FUNCTION_BLOCK ActuatorBaseExt (* Composite Function Block Type *)
  (* Standard: 61499-2 *)
  (* Version 1.0.1, 10/17/2023, ApplicationLibDevTeam, Schneider Electric, First Version *)
  PACKAGE Flexbridge.FestoMPS400;
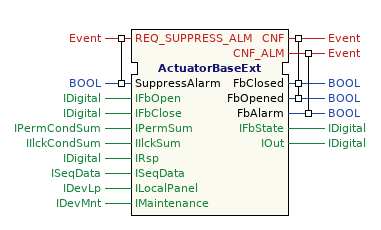
  EVENT_INPUT
    REQ_SUPPRESS_ALM WITH SuppressAlarm; (* Request to update the alarm suppress status *)
  END_EVENT
  EVENT_OUTPUT
    CNF WITH FbClosed, FbOpened; (* Execution confirmation *)
    CNF_ALM WITH FbAlarm; (* Execution confirmation of alarm *)
  END_EVENT
  VAR_INPUT
    SuppressAlarm : BOOL; (* 1 = Suppress alarm in HMI *)
  END_VAR
  VAR_OUTPUT
    FbClosed : BOOL; (* 1 = Closed *)
    FbOpened : BOOL; (* 1 = Opened *)
    FbAlarm : BOOL; (* 1 = Feedback failure alarm is active *)
  END_VAR
  SOCKETS
    IFbOpen : IDigital; (* Open feedback signal adapter *)
    IFbClose : IDigital; (* Close feedback signal adapter *)
    IPermSum : IPermCondSum(DeviceType := UniDirectional, ServiceState := TRUE); (* Permission condition summary chain input from permcondsum block *)
    IIlckSum : IIlckCondSum(DeviceType := UniDirectional, ServiceState := TRUE); (* Interlock condition summary chain input from ilckcondsum block *)
  END_SOCKETS
  SOCKETS
    IRsp : IDigital; (* Program remote setpoint interface adapter *)
    ISeqData : ISeqData; (* Sequence control interface adapter, Controls the block when owner is in program local *)
    ILocalPanel : IDevLp; (* Local panel Interface adapter *)
    IMaintenance : IDevMnt; (* Maintenance data Interface adapter *)
  END_SOCKETS
  PLUGS
    IFbState : IDigital; (* Current feedback status Interface adapter *)
    IOut : IDigital; (* Current Output status Interface adapter *)
  END_PLUGS
  (* Control *)
  (* Permissive *)
  (* Interlock *)
  (* Input Hardware Interface *)
  (* Service Connection *)
  (* Output Interface *)
  (* Hardware Output Interface *)
  FBS
    serviceManager : ValveServiceManager;
    fbConv : intToBool; {SET_ATTRIBUTE(Configuration.Component.HideUnusedPorts, )}
    actuatorBase : ActuatorBase; {SET_ATTRIBUTE(Configuration.Component.HideUnusedPorts, )}
  END_FBS
  EVENT_CONNECTIONS
    actuatorBase.CNF_FB_STS TO CNF;
    REQ_SUPPRESS_ALM TO actuatorBase.REQ_SUPPRESS_ALM;
    IPermSum.PERM_IND TO actuatorBase.REQ_PERM;
    IIlckSum.COND_IND TO actuatorBase.REQ_ILCK;
    actuatorBase.CNF_FB_STS TO IFbState.REQ;
    actuatorBase.CNF_MODE TO IIlckSum.REQ;
    actuatorBase.CNF_OUT TO IOut.REQ;
    actuatorBase.CNF_FB_ALM TO CNF_ALM;
    actuatorBase.CNF_ALM TO IFbState.REQ_STATUS;
    IPermSum.CHECK_SERVICE TO IPermSum.CNF_SERVICE;
    IIlckSum.CHECK_SERVICE TO IIlckSum.CNF_SERVICE;
    actuatorBase.CNF_MODE TO IOut.REQ_STATUS;
    IFbOpen.REQ TO fbConv.REQ1;
    fbConv.CNF1 TO actuatorBase.REQ_FB;
    IFbClose.REQ TO fbConv.REQ2;
    fbConv.CNF2 TO actuatorBase.REQ_FB;
    actuatorBase.CNF_OWNER TO IIlckSum.REQ_OWNER;
  END_CONNECTIONS
  DATA_CONNECTIONS
    actuatorBase.FbAlarm TO FbAlarm;
    IIlckSum.CondType TO actuatorBase.IlckType;
    IIlckSum.CondPos TO actuatorBase.IlckPos;
    actuatorBase.FbStatus TO IFbState.Value;
    actuatorBase.AlarmStatus TO IFbState.Status;
    actuatorBase.Maintenance TO IIlckSum.Suppress;
    IPermSum.PermPassive TO actuatorBase.PermClose;
    actuatorBase.FbOpened TO FbOpened;
    actuatorBase.FbClosed TO FbClosed;
    IIlckSum.State TO actuatorBase.IlckCond;
    actuatorBase.Out TO IOut.Value;
    actuatorBase.Simulation TO IOut.Status;
    IPermSum.PermActive1 TO actuatorBase.PermOpen;
    IFbOpen.Value TO fbConv.IN1;
    IFbClose.Value TO fbConv.IN2;
    fbConv.OUT1 TO actuatorBase.FbOpen;
    fbConv.OUT2 TO actuatorBase.FbClose;
    SuppressAlarm TO actuatorBase.SuppressAlarm;
    actuatorBase.CurrentOwner TO IIlckSum.CurrentOwner;
  END_CONNECTIONS
  ADAPTER_CONNECTIONS
    IMaintenance TO serviceManager.IMaint;
    ILocalPanel TO serviceManager.28;
    ISeqData TO serviceManager.31;
    serviceManager.14 TO actuatorBase.187;
    IRsp TO serviceManager.IRsp;
  END_CONNECTIONS
END_FUNCTION_BLOCK
